(* PLC project Vn_fb_ftrig, Beckhoff Automation GmbH TwinCAT PLC Control 3.5.13.21 *)
(* stored: creationDateTime 1970-01-01T00:00:00 *)

PROGRAM Vn_fb_ftrig

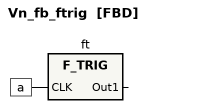
(* FBD diagram, written out as Structured Text *)
ft(CLK := a);
END_PROGRAM
